FUNCTION_BLOCK FB_ValveMonitor (* Migrated from IEC 61131-3 ST *)
  (* Standard: 61499-2 *)
  (* Version 1.0, 2026-11-06, st2fb *)
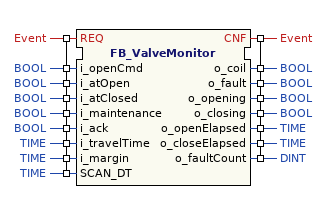
  EVENT_INPUT
    REQ WITH i_openCmd, i_atOpen, i_atClosed, i_maintenance, i_ack, i_travelTime, i_margin, SCAN_DT;
  END_EVENT
  EVENT_OUTPUT
    CNF WITH o_coil, o_fault, o_opening, o_closing, o_openElapsed, o_closeElapsed, o_faultCount;
  END_EVENT
  VAR_INPUT
    i_openCmd : BOOL;
    i_atOpen : BOOL;
    i_atClosed : BOOL;
    i_maintenance : BOOL;
    i_ack : BOOL;
    i_travelTime : TIME;
    i_margin : TIME;
    SCAN_DT : TIME;
  END_VAR
  VAR_OUTPUT
    o_coil : BOOL;
    o_fault : BOOL;
    o_opening : BOOL;
    o_closing : BOOL;
    o_openElapsed : TIME;
    o_closeElapsed : TIME;
    o_faultCount : DINT;
  END_VAR
  VAR
    ST2FB_NOW : TIME := T#0s;
    statOpenBudget : TIME := T#0s;
    statCloseBudget : TIME := T#0s;
    tempBudget : TIME := T#0s;
    OT_IN : BOOL := FALSE;
    OT_PT : TIME := T#0s;
    OT_Q : BOOL := FALSE;
    OT_ET : TIME := T#0s;
    OT_STATE : INT := 0;
    OT_PREV_IN : BOOL := FALSE;
    OT_START_TIME : TIME := T#0s;
    CT_IN : BOOL := FALSE;
    CT_PT : TIME := T#0s;
    CT_Q : BOOL := FALSE;
    CT_ET : TIME := T#0s;
    CT_STATE : INT := 0;
    CT_PREV_IN : BOOL := FALSE;
    CT_START_TIME : TIME := T#0s;
    FE_CLK : BOOL := FALSE;
    FE_Q : BOOL := FALSE;
    FE_M : BOOL := FALSE;
  END_VAR
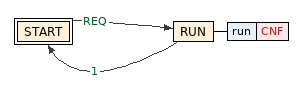
  EC_STATES
    START;
    RUN : run -> CNF;
  END_STATES
  EC_TRANSITIONS
    START TO RUN := REQ;
    RUN TO START := 1;
  END_TRANSITIONS
  ALGORITHM run IN ST:
ST2FB_NOW := ST2FB_NOW + SCAN_DT;
IF NOT i_maintenance THEN
  tempBudget := i_travelTime + i_margin;
  o_coil := i_openCmd AND NOT o_fault;
  IF NOT o_opening THEN
    statOpenBudget := tempBudget;
  END_IF;
  IF NOT o_closing THEN
    statCloseBudget := tempBudget;
  END_IF;
  o_opening := o_coil AND NOT i_atOpen;
  o_closing := NOT o_coil AND NOT i_atClosed;

  OT_IN := o_opening;
  OT_PT := statOpenBudget;
  IF (OT_STATE = 0) AND NOT OT_PREV_IN AND OT_IN THEN
    OT_STATE := 1;
    OT_Q := FALSE;
    OT_START_TIME := ST2FB_NOW;
  ELSE
    IF NOT OT_IN THEN
      OT_ET := T#0s;
      OT_Q := FALSE;
      OT_STATE := 0;
    ELSIF OT_STATE = 1 THEN
      IF OT_START_TIME + OT_PT <= ST2FB_NOW THEN
        OT_STATE := 2;
        OT_Q := TRUE;
        OT_ET := OT_PT;
      ELSE
        OT_ET := ST2FB_NOW - OT_START_TIME;
      END_IF;
    END_IF;
  END_IF;
  OT_PREV_IN := OT_IN;
  o_openElapsed := OT_ET;

  CT_IN := o_closing;
  CT_PT := statCloseBudget;
  IF (CT_STATE = 0) AND NOT CT_PREV_IN AND CT_IN THEN
    CT_STATE := 1;
    CT_Q := FALSE;
    CT_START_TIME := ST2FB_NOW;
  ELSE
    IF NOT CT_IN THEN
      CT_ET := T#0s;
      CT_Q := FALSE;
      CT_STATE := 0;
    ELSIF CT_STATE = 1 THEN
      IF CT_START_TIME + CT_PT <= ST2FB_NOW THEN
        CT_STATE := 2;
        CT_Q := TRUE;
        CT_ET := CT_PT;
      ELSE
        CT_ET := ST2FB_NOW - CT_START_TIME;
      END_IF;
    END_IF;
  END_IF;
  CT_PREV_IN := CT_IN;
  o_closeElapsed := CT_ET;

  IF i_ack THEN
    o_fault := FALSE;
  ELSIF OT_Q OR CT_Q OR (i_atOpen AND i_atClosed) THEN
    o_fault := TRUE;
  END_IF;
  FE_CLK := o_fault;
  FE_Q := FE_CLK AND NOT FE_M;
  FE_M := FE_CLK;
  IF FE_Q THEN
    o_faultCount := o_faultCount + 1;
  END_IF;
END_IF;
  END_ALGORITHM
END_FUNCTION_BLOCK
